Fanuc KAREL source: KT00729.KL

PROGRAM KT00729
%NOLOCKGROUP
VAR
  C1: CONFIG
  C2: CONFIG
  OUT: INTEGER
BEGIN
  C1.CFG_FLIP = TRUE
  C2.CFG_FLIP = FALSE
  C1.CFG_FLIP = TRUE
  C2.CFG_FLIP = FALSE
  OUT = ARRAY_LEN(C1)
END KT00729
